// TIA Portal V20 export
// export: Created 2026-10-20T18:55:50.8044859Z, ExportSetting None, DisplayName Totally Integrated Automation Portal, DisplayVersion V20 Update 6, DisplayName TIA Portal Openness, DisplayVersion V20 Update 6, DisplayName TIA Portal Version Control Interface, DisplayVersion V20 Update 6, DisplayName SINAMICS Startdrive Advanced, DisplayVersion V20 SP1, DisplayName SINAMICS Startdrive G130, G150, S120, S150, SINAMICS MV, G220, S200, S210, DisplayVersion V20 SP1, DisplayName SINAMICS Startdrive G110M, G120, G120C, G120D, G120P, G115D, DisplayVersion V20 SP1, DisplayName STEP 7 Professional, DisplayVersion V20 Update 6, DisplayName STEP 7 Safety, DisplayVersion V20 Update 2, DisplayName WinCC Basic/Comfort/Advanced, DisplayVersion V20 Update 6, DisplayName WinCC Unified, DisplayVersion V20 Update 6
VAR_GLOBAL   // PLC tag table "Lock_6"
   "Solenoid Enable_6" AT %Q1377.0 : Bool;
   Lock_6_Estop_CH1 AT %I1798.2 : Bool;
   Lamps_6 AT %QB1376 : Byte;
   "Lock Reset_6" AT %Q1490.0 : Bool;
   Lock_6_Estop_CH2 AT %I1798.3 : Bool;
   Lock_6_Closed_CH1 AT %I1798.0 : Bool;
   Lock_6_Closed_CH2 AT %I1798.1 : Bool;
   Switches_6 AT %IB1280 : Byte;
   Lock_6_Reset_Input1 AT %Q1799.0 : Bool;
   Lock_6_Reset_Input2 AT %Q1799.1 : Bool;
   Lock_6_Reset_Input3 AT %Q1799.2 : Bool;
   Lock_6_Reset_Input4 AT %Q1799.3 : Bool;
   "Lock Position_6" AT %I1342.0 : Bool;
   "Guard Position_6" AT %I1341.0 : Bool;
END_VAR
